FUNCTION_BLOCK ProcessingSequence1 (* Composite Function Block Type *)
  (* Standard: 61499-2 *)
  (* Version 0.0, 7/2/2026, template *)
  PACKAGE Main;
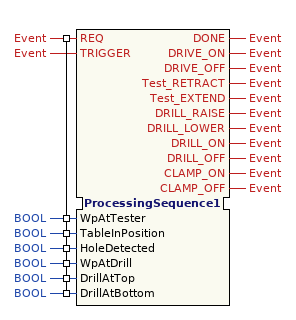
  EVENT_INPUT
    REQ WITH WpAtTester, TableInPosition, HoleDetected, WpAtDrill, DrillAtTop, DrillAtBottom; (* Normal Execution Request *)
    TRIGGER;
  END_EVENT
  EVENT_OUTPUT
    DONE; (* Initialization Confirm *)
    DRIVE_ON; (* Execution Confirmation *)
    DRIVE_OFF;
    Test_RETRACT;
    Test_EXTEND;
    DRILL_RAISE;
    DRILL_LOWER;
    DRILL_ON;
    DRILL_OFF;
    CLAMP_ON;
    CLAMP_OFF;
  END_EVENT
  VAR_INPUT
    WpAtTester : BOOL; (* Input event qualifier *)
    TableInPosition : BOOL;
    HoleDetected : BOOL;
    WpAtDrill : BOOL;
    DrillAtTop : BOOL;
    DrillAtBottom : BOOL;
  END_VAR
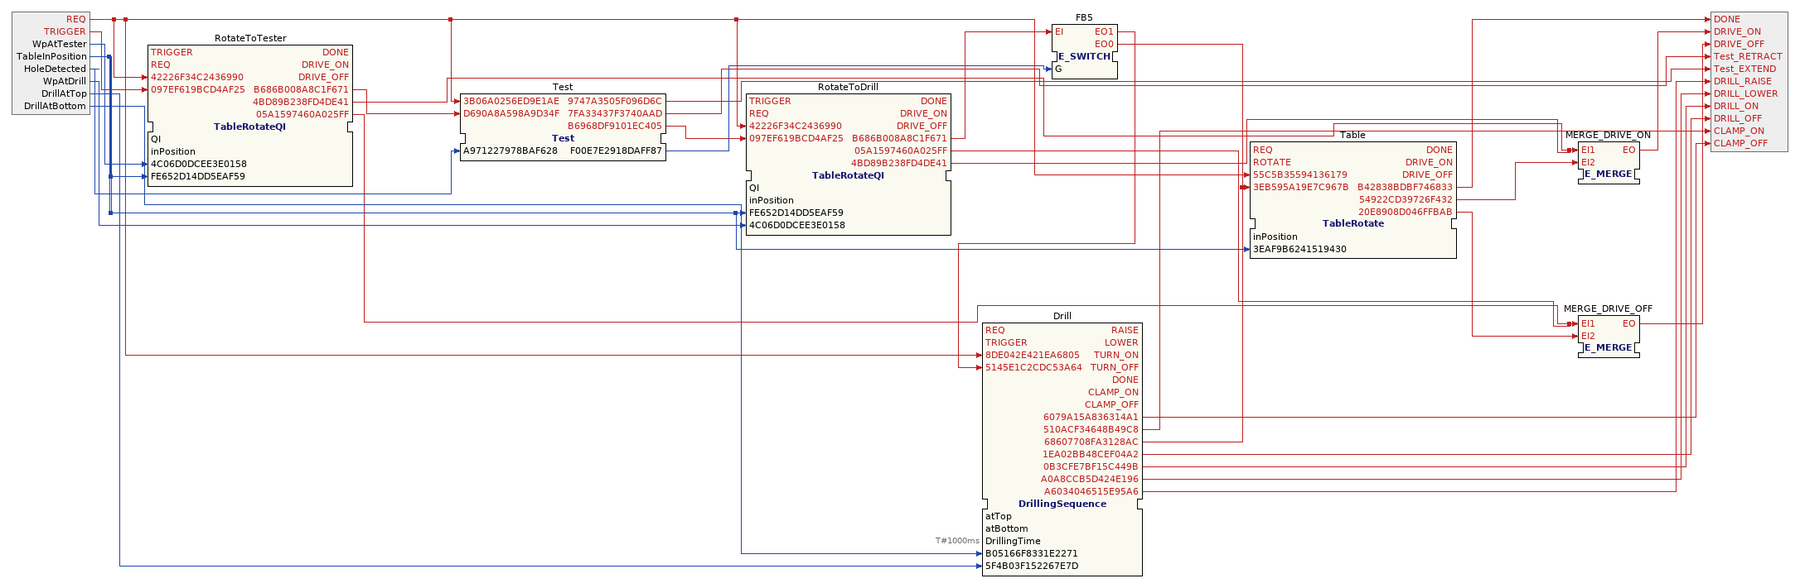
  FBS
    RotateToTester : TableRotateQI;
    Test : Test;
    RotateToDrill : TableRotateQI;
    Drill : DrillingSequence(DrillingTime := T#1000ms);
    FB5 : E_SWITCH;
    Table : TableRotate;
    MERGE_DRIVE_ON : E_MERGE;
    MERGE_DRIVE_OFF : E_MERGE;
  END_FBS
  EVENT_CONNECTIONS
    MERGE_DRIVE_OFF.EO TO DRIVE_OFF;
    MERGE_DRIVE_ON.EO TO DRIVE_ON;
    REQ TO RotateToTester.42226F34C2436990;
    REQ TO Test.3B06A0256ED9E1AE;
    REQ TO Drill.8DE042E421EA6805;
    REQ TO RotateToDrill.42226F34C2436990;
    REQ TO Table.55C5B35594136179;
    TRIGGER TO RotateToTester.097EF619BCD4AF25;
    RotateToTester.B686B008A8C1F671 TO Test.D690A8A598A9D34F;
    RotateToTester.4BD89B238FD4DE41 TO MERGE_DRIVE_ON.EI1;
    RotateToTester.05A1597460A025FF TO MERGE_DRIVE_OFF.EI1;
    Table.B42838BDBF746833 TO DONE;
    Drill.6079A15A836314A1 TO CLAMP_OFF;
    Drill.510ACF34648B49C8 TO CLAMP_ON;
    Drill.68607708FA3128AC TO Table.3EB595A19E7C967B;
    Drill.1EA02BB48CEF04A2 TO DRILL_OFF;
    Drill.0B3CFE7BF15C449B TO DRILL_ON;
    Drill.A0A8CCB5D424E196 TO DRILL_LOWER;
    Drill.A6034046515E95A6 TO DRILL_RAISE;
    Test.9747A3505F096D6C TO Test_EXTEND;
    Test.7FA33437F3740AAD TO Test_RETRACT;
    RotateToDrill.B686B008A8C1F671 TO FB5.EI;
    FB5.EO1 TO Drill.5145E1C2CDC53A64;
    Test.B6968DF9101EC405 TO RotateToDrill.097EF619BCD4AF25;
    RotateToDrill.05A1597460A025FF TO MERGE_DRIVE_OFF.EI1;
    RotateToDrill.4BD89B238FD4DE41 TO MERGE_DRIVE_ON.EI1;
    Table.54922CD39726F432 TO MERGE_DRIVE_ON.EI2;
    Table.20E8908D046FFBAB TO MERGE_DRIVE_OFF.EI2;
    FB5.EO0 TO Table.3EB595A19E7C967B;
  END_CONNECTIONS
  DATA_CONNECTIONS
    WpAtTester TO RotateToTester.4C06D0DCEE3E0158;
    TableInPosition TO RotateToTester.FE652D14DD5EAF59;
    TableInPosition TO RotateToDrill.FE652D14DD5EAF59;
    TableInPosition TO Table.3EAF9B6241519430;
    WpAtDrill TO RotateToDrill.4C06D0DCEE3E0158;
    HoleDetected TO Test.A971227978BAF628;
    Test.F00E7E2918DAFF87 TO FB5.G;
    DrillAtBottom TO Drill.B05166F8331E2271;
    DrillAtTop TO Drill.5F4B03F152267E7D;
  END_CONNECTIONS
END_FUNCTION_BLOCK
